(* IEC 61131-3 sources: ConveyorControl-with-PLC/4E_Gruppe1_Graf_Projekt1_HMI/Network/LseRtkAlarm, 1 file *)

(* ---- ONE_LseRtkAlarm_Table.st ---- *)
#define OBJECTS_CONFIG

#include "..\..\Class\_AlarmX0Para\_AlarmX0Para.h"
#include <.\lsl_st_mt.h>
#include "..\..\Class\_AlarmXBuffer\AlarmXBuffer.h"

FUNCTION GLOBAL TAB ONE_LseRtkAlarm
-1$UINT, 0$UINT,
0$UINT, 0$UINT,

7$UDINT,
TO_UDINT(1738954212), "_AlarmDisplay", 0$UINT, 7$UINT, 2$UINT,
TO_UDINT(800276940), "_AlarmX0Para", 0$UINT, 7$UINT, 1$UINT,
TO_UDINT(315844732), "_AlarmX1Para", 0$UINT, 2$UINT, 1$UINT,
TO_UDINT(2835625764), "_AlarmXBuffer", 0$UINT, 14$UINT, 1$UINT,
TO_UDINT(3509550928), "_HotAlarm", 0$UINT, 1$UINT, 1$UINT,
TO_UDINT(2980745877), "_MyIO", 0$UINT, 3$UINT, 0$UINT,
TO_UDINT(3043040051), "_ScrollArea", 0$UINT, 14$UINT, 0$UINT,

_NO_ATTR, TO_UDINT(378942885), "ALARMHISTORY",
_NO_ATTR, TO_UDINT(4248743175), "ALARMTEMPORARY",

_NO_ATTR, TO_UDINT(3323358457), "EMERGENCYSTOP",

_NO_ATTR, TO_UDINT(108736354), "SERVERERROR",

_NO_ATTR, TO_UDINT(3212185425), "_ALARMXBUFFER1",

_NO_ATTR, TO_UDINT(4293868080), "HOTALARM",

//Internal connections
0$UDINT,
0$UDINT,
0$UDINT,
0$UDINT,

//Initialization values
0$UDINT,
15$UDINT,
TO_UDINT(0), "VerticalLevel", TO_UDINT(1),//|LseRtkAlarm.AlarmHistory.VerticalLevel;
TO_UDINT(0), "LineWidth", TO_UDINT(1),//|LseRtkAlarm.AlarmHistory.LineWidth;
TO_UDINT(0), "ExtendedScrollBar", TO_UDINT(0),//|LseRtkAlarm.AlarmHistory.ExtendedScrollBar;
TO_UDINT(0), "HistoryTemporary", TO_UDINT(0),//|LseRtkAlarm.AlarmHistory.HistoryTemporary;
TO_UDINT(0), "MaxNo", TO_UDINT(100),//|LseRtkAlarm.AlarmHistory.MaxNo;
TO_UDINT(0), "Filter", TO_UDINT(0),//|LseRtkAlarm.AlarmHistory.Filter;
TO_UDINT(1), "VerticalLevel", TO_UDINT(1),//|LseRtkAlarm.AlarmTemporary.VerticalLevel;
TO_UDINT(1), "LineWidth", TO_UDINT(1),//|LseRtkAlarm.AlarmTemporary.LineWidth;
TO_UDINT(1), "ExtendedScrollBar", TO_UDINT(0),//|LseRtkAlarm.AlarmTemporary.ExtendedScrollBar;
TO_UDINT(1), "HistoryTemporary", TO_UDINT(1),//|LseRtkAlarm.AlarmTemporary.HistoryTemporary;
TO_UDINT(1), "MaxNo", TO_UDINT(100),//|LseRtkAlarm.AlarmTemporary.MaxNo;
TO_UDINT(1), "Filter", TO_UDINT(10),//|LseRtkAlarm.AlarmTemporary.Filter;
TO_UDINT(2), "Config", TO_UDINT(1),//|LseRtkAlarm.EmergencyStop.Config;
TO_UDINT(3), "Config", TO_UDINT(2),//|LseRtkAlarm.ServerError.Config;
TO_UDINT(4), "No", TO_UDINT(64),//|LseRtkAlarm._AlarmXBuffer1.No;

//Symbolic initialization values
0$UDINT,
0$UDINT,

//Initialization of string values
0$UDINT,
0$UDINT,

//Configuration of tasks (RealTime, Cyclic, Background)
0$UDINT,
0$UDINT,

0$UDINT,
0$UDINT,

0$UDINT,
0$UDINT,

//External connections
0$UDINT,
3$UDINT,
TO_UDINT(0), "Lse", C_DIR, TO_UDINT(299963966), "Lse","Lse",
TO_UDINT(1), "Lse", C_DIR, TO_UDINT(299963966), "Lse","Lse",
TO_UDINT(5), "Lse", C_DIR, TO_UDINT(299963966), "Lse","Lse",

//Magic internal connections
0$UDINT,
0$UDINT,

//Configuration of timeslots of tasks (RealTime, Cyclic)
#ifdef __LSLLDR_TIMESLOTS__
0$UDINT,
0$UDINT,

0$UDINT,
0$UDINT,

#endif //__LSLLDR_TIMESLOTS__

//MultiMaster connections
#ifdef __LSLLDR_MULTIMASTER__
0$UDINT,
0$UDINT,
#endif //__LSLLDR_MULTIMASTER__

END_FUNCTION
